PROGRAM main
  VAR
    NGFel : BOOL;
    NGLe : BOOL;
    Vegallas_fent : BOOL;
    Vegallas_lent : BOOL;
    Kapu_fel : BOOL;
    Allj : BOOL;
    Kapu_le : BOOL;
    Lampa : BOOL;
    Time_limit : TIME := T#5s;
    RealTime : TIME;
    Timer_on : BOOL;
    Time_contivnue : BOOL;
    TON0 : TON;
  END_VAR
  VAR  (* added by the conversion: wires and edge detectors of the diagram *)
    _EQ3_ENO : BOOL;
    _EQ3_OUT : BOOL;
    _EQ15_ENO : BOOL;
    _EQ15_OUT : BOOL;
  END_VAR

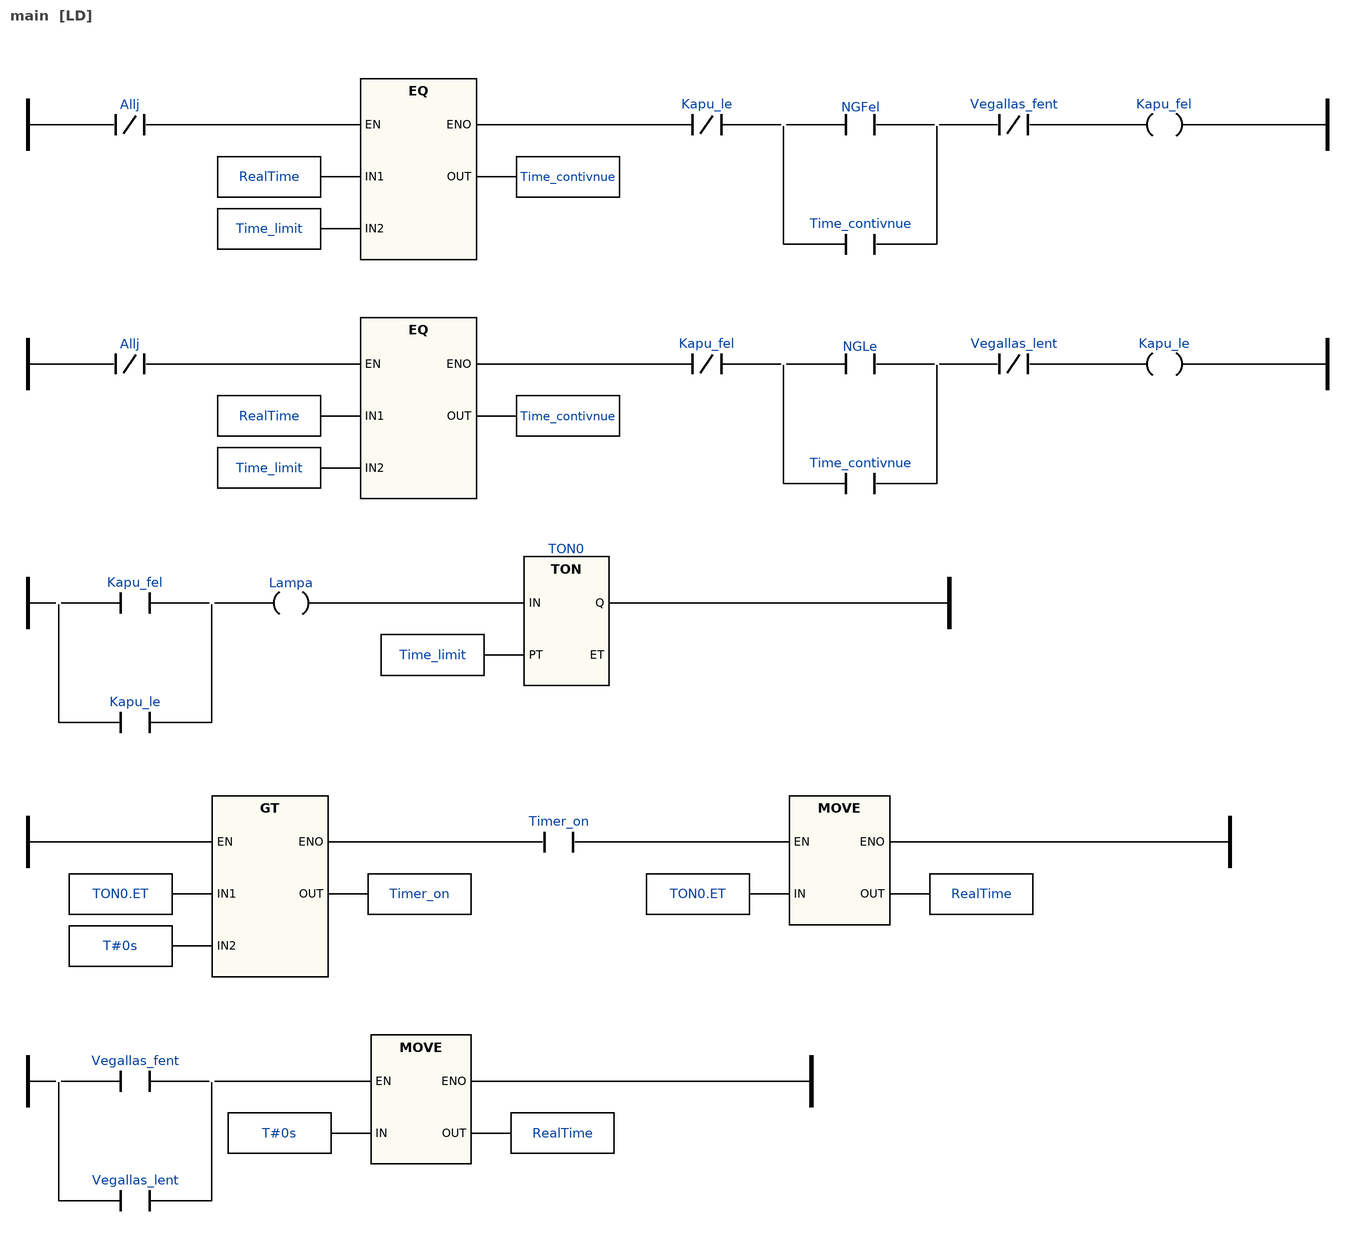
(* LD diagram, written out as Structured Text *)
_EQ3_OUT := EQ(EN := NOT Allj, IN1 := RealTime, IN2 := Time_limit, ENO => _EQ3_ENO);
Kapu_fel := _EQ3_ENO AND NOT Kapu_le AND (NGFel OR Time_contivnue) AND NOT Vegallas_fent;
IF _EQ3_ENO THEN Time_contivnue := _EQ3_OUT; END_IF;
_EQ15_OUT := EQ(EN := NOT Allj, IN1 := RealTime, IN2 := Time_limit, ENO => _EQ15_ENO);
Kapu_le := _EQ15_ENO AND NOT Kapu_fel AND (NGLe OR Time_contivnue) AND NOT Vegallas_lent;
IF _EQ15_ENO THEN Time_contivnue := _EQ15_OUT; END_IF;
Lampa := Kapu_fel OR Kapu_le;
Timer_on := TON0.ET > T#0s;
IF Timer_on THEN RealTime := TON0.ET; END_IF;
IF Vegallas_fent OR Vegallas_lent THEN RealTime := T#0s; END_IF;
TON0(IN := Kapu_fel OR Kapu_le, PT := Time_limit);
END_PROGRAM
